Universal Robots PolyScope program: Weight_detection.urp

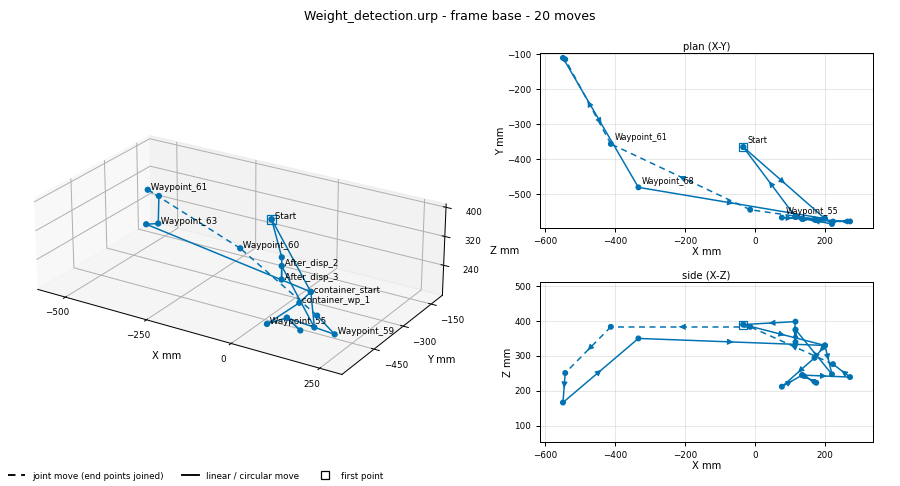
[picture p0: tool path of Weight_detection.urp in frame base, 20 of 20 moves have a stored position in this frame; points joined in program order, loops and branches not executed]
Program Weight_detection (installation=default directory=/programs/02 Main Routines createdIn=5.19.0 lastSavedIn=5.19.0 robotSerialNumber=20245590068)
Calibrated DH parameters: a=[0.00013, -0.03651, -0.389144, 0.000102, 0.000008, 0]; d=[0.162613, 192.230671, -179.915756, -12.181517, 0.099698, 0.099535]; alpha=[1.57038, 0.002205, 0.004138, 1.570804, -1.571025, 0]; deltaTheta=[-0.000001, 1.484886, 4.928506, -0.130209, 0, 0]
InitVariablesNode
Robot Program (runOnlyOnce=true)
  Folder powder dispensing variable init
    Start_thread := False
    kp := 0.0005
    ki := 0.002
    kd := 0.02
    dt := 0.05
    Weight_value := get_weight()
    Target_weight :=  (valueSource=Operator message=Enter the Target weight to be dispensed in gm valueType=Float)
    Integral_error := 0
    current_error := 0
    previous_error := 0
    tilt_increment := 0
    tilt_angle := -1
  Script file /programs/04 Scripts/Weight_scale_socket.script
    | def get_weight():
    | 	socket_open("192.168.12.190", 3002)
    | 	textmsg("socket opened successfully!")
    | 	socket_send_string("GET_WEIGHT")
    | 	sync()
    | 	sleep(0.5)
    | 	receiveFromServ = socket_read_ascii_float(6)
    | 	while (receiveFromServ[0] <1):
    | 		sleep(0.5)
    | 		receiveFromServ = socket_read_ascii_float(1)
    | 		textmsg("retrying read:", receiveFromServ)
    | 	end
    | 	textmsg("Received weight:", receiveFromServ[1])
    | 	socket_close()
    | 	return receiveFromServ[1]
    | end
  Script file /programs/04 Scripts/dosing_pid.script
    | def dosing_pid(Target_weight):
    | 	#kp = 0.005
    | 	#ki = 0.02
    | 	#kd = 0.2
    | 	#dt = 0.05
    | 	#current_error = 0.0
    | 	#Integral_error = 0.0
    | 	#previous_error = 0.0
    | 	#tilt_angle = -1.0
    | 	max_tilt_angle = -0.55
    | 	#current_pose = get_actual_tcp_pose()
    | 
    | 	while ( Weight_value < Target_weight and tilt_angle < max_tilt_angle):
    | 		Weight_value = get_weight()
    | 		current_error = Target_weight - Weight_value
    | 		Integral_error = Integral_error + current_error*dt
    | 		derivative = (current_error - previous_error) / dt
    | 		tilt_increment = (kp * current_error) + (ki * Integral_error) + (kd * derivative)
    | 		current_pose = get_actual_tcp_pose()
    | 		tilt_angle = current_pose[4]
    | 		new_pose = pose_trans(current_pose, p[(tilt_increment/5), 0, 0, 0, tilt_increment, 0])
    | 		movel(new_pose, a = 0.075, v = 0.025, t = 0, r = 0)
    | 		previous_error = current_error
    | 		sleep(dt)
    | 	end
    | end
  MoveL speed 250 mm/s, acceleration 1200 mm/s^2 (useActiveTCP=true) feature=Base
    Waypoint Start: TCP in base x=-33.065 y=-365.399 z=389.873 mm, rx=0 ry=0 rz=2.7258 rad; joints [-73.774, -70.638, -96.716, -102.629, 90.121, 40.001] deg; TCP offset x=0 y=0 z=161 mm, rx=3.1415 ry=0 rz=0 rad
  SuppressedNode
    MoveL speed 50 mm/s, acceleration 300 mm/s^2 (useActiveTCP=true) feature=Base
      Waypoint Waypoint_53: motionParameters(jointSpeed=1.047198 jointAcceleration=1.396263 cartesianSpeed=0.1 cartesianAcceleration=0.3); TCP in base x=200.65 y=-570.239 z=330.084 mm, rx=1.3605 ry=0.0217 rz=2.6816 rad; joints [-43.952, -124.342, -49.589, -141.868, 58.423, 68.107] deg
      Waypoint Waypoint_54: motionParameters(jointSpeed=1.047198 jointAcceleration=1.396263 cartesianSpeed=0.05 cartesianAcceleration=0.3); TCP in base x=170.614 y=-572.151 z=294.509 mm, rx=1.2595 ry=-0.0083 rz=2.7877 rad; joints [-46.577, -118.755, -62.143, -128.361, 58.907, 59.792] deg
      Loop Counting (count=3) loopVariable(name=Loop_4)
        Waypoint Waypoint_55: motionParameters(jointSpeed=1.047198 jointAcceleration=1.396263 cartesianSpeed=0.05 cartesianAcceleration=0.3); TCP in base x=77.281 y=-567.309 z=212.068 mm, rx=1.2595 ry=-0.0083 rz=2.7877 rad; joints [-52.608, -113.129, -83.31, -109.754, 55.252, 54.186] deg
          Until TOOL_CONTACT_DETECTION (allowActions=false retraction=0 decelerationAcceleration=3 decelerationAngularAcceleration=34.906585)
        Waypoint Waypoint_56: motionParameters(jointSpeed=1.047198 jointAcceleration=1.396263 cartesianSpeed=0.05 cartesianAcceleration=0.3); TCP in base x=135.568 y=-570.868 z=245.215 mm, rx=1.4769 ry=-0.0183 rz=2.6796 rad; joints [-47.325, -120.782, -69.397, -128.377, 54.155, 64.498] deg
      Loop Counting (count=2) loopVariable(name=Loop_5)
        Waypoint Waypoint_1: motionParameters(jointSpeed=1.047198 jointAcceleration=1.396263 cartesianSpeed=0.4 cartesianAcceleration=1.2); TCP in base x=175.61 y=-574.617 z=223.224 mm, rx=1.7438 ry=-0.031 rz=2.516 rad; joints [-43.942, -131.598, -59.719, -142.336, 52.9, 75.006] deg
        Waypoint Waypoint_56: motionParameters(jointSpeed=1.047198 jointAcceleration=1.396263 cartesianSpeed=0.05 cartesianAcceleration=0.3); TCP in base x=135.568 y=-570.868 z=245.215 mm, rx=1.4769 ry=-0.0183 rz=2.6796 rad; joints [-47.325, -120.782, -69.397, -128.377, 54.155, 64.498] deg
      Waypoint Waypoint_59: motionParameters(jointSpeed=1.047198 jointAcceleration=1.396263 cartesianSpeed=0.05 cartesianAcceleration=0.3); TCP in base x=272.401 y=-578.183 z=239.561 mm, rx=2.127 ry=0.1139 rz=2.1556 rad; joints [-37.816, -154.733, -25.502, -178.522, 53.445, 96.624] deg
      Waypoint Waypoint_58: motionParameters(jointSpeed=1.047198 jointAcceleration=1.396263 cartesianSpeed=0.05 cartesianAcceleration=0.3); TCP in base x=223.649 y=-578.478 z=276.546 mm, rx=2.1743 ry=-0.0441 rz=2.0587 rad; joints [-41.771, -153.265, -25.455, -184.54, 55.381, 96.631] deg
  SuppressedNode
    MoveJ speed 30 deg/s, acceleration 50 deg/s^2 (useActiveTCP=true) feature=Base
      Waypoint Waypoint_60: motionParameters(jointSpeed=0.349066 jointAcceleration=0.523599 cartesianSpeed=0.25 cartesianAcceleration=1.2 blendRadius=0.05); TCP in base x=-13.316 y=-544.772 z=383.372 mm, rx=2.2082 ry=0.0375 rz=2.0976 rad; joints [-53.447, -120.321, -68.514, -175.377, 39.556, 98.101] deg
      Waypoint Waypoint_61: motionParameters(jointSpeed=0.349066 jointAcceleration=0.523599 cartesianSpeed=0.25 cartesianAcceleration=1.2 blendRadius=0.05); TCP in base x=-412.189 y=-356.447 z=383.372 mm, rx=1.7517 ry=-0.74 rz=1.6007 rad; joints [-101.195, -120.321, -68.514, -175.377, 39.556, 98.101] deg
      Waypoint Waypoint_62: motionParameters(jointSpeed=0.349066 jointAcceleration=0.523599 cartesianSpeed=0.25 cartesianAcceleration=1.2); TCP in base x=-542.659 y=-114.282 z=251.262 mm, rx=1.813 ry=-0.6794 rz=1.6553 rad; joints [-123.661, -111.262, -103.952, -159.22, 12.548, 108.767] deg
  SuppressedNode
    MoveL speed 250 mm/s, acceleration 1200 mm/s^2 (useActiveTCP=true) feature=Base
      Waypoint Waypoint_63: motionParameters(jointSpeed=1.047198 jointAcceleration=1.396263 cartesianSpeed=0.05 cartesianAcceleration=0.3); TCP in base x=-532.496 y=-127.81 z=184.034 mm, rx=1.813 ry=-0.6794 rz=1.6553 rad; joints [-121.653, -117.001, -107.545, -147.984, 14.526, 106.805] deg
      If Target_weight<Weight_value (checkContinuously=true)
        Script: dosing_pid()
      Waypoint Waypoint_64: motionParameters(jointSpeed=1.047198 jointAcceleration=1.396263 cartesianSpeed=0.05 cartesianAcceleration=0.3); TCP in base x=-576.035 y=-66.27 z=306.74 mm, rx=0.8621 ry=-0.2554 rz=2.1952 rad; joints [-142.141, -87.685, -107.535, -64.498, 50.077, -8.596] deg
      Waypoint Waypoint_65: motionParameters(jointSpeed=1.047198 jointAcceleration=1.396263 cartesianSpeed=0.05 cartesianAcceleration=0.3); TCP in base x=-581.965 y=-59.291 z=312.082 mm, rx=0.8621 ry=-0.2554 rz=2.1952 rad; joints [-143.275, -88.018, -106.65, -64.116, 50.29, -10.05] deg
      Waypoint Waypoint_66: motionParameters(jointSpeed=1.047198 jointAcceleration=1.396263 cartesianSpeed=0.5 cartesianAcceleration=1.2); TCP in base x=-581.965 y=-59.291 z=290.576 mm, rx=0.8621 ry=-0.2554 rz=2.1952 rad; joints [-143.281, -88.87, -109.094, -60.824, 50.286, -10.043] deg
      Waypoint Waypoint_67: TCP in base x=-581.965 y=-59.291 z=350.142 mm, rx=1.7575 ry=-0.6778 rz=1.6965 rad; joints [-131.863, -101.687, -97.87, -162.913, 4.302, 96.426] deg
  SuppressedNode
    MoveJ speed 60 deg/s, acceleration 80 deg/s^2 (useActiveTCP=true) feature=Base
      Waypoint Waypoint_68: motionParameters(jointSpeed=1.047198 jointAcceleration=1.396263 cartesianSpeed=0.25 cartesianAcceleration=1.2); TCP in base x=-333.293 y=-480.744 z=350.142 mm, rx=2.2175 ry=0.1409 rz=2.2091 rad; joints [-82.414, -101.687, -97.87, -162.913, 4.302, 96.426] deg
  Folder powder dispensing
    Loop While (checkContinuously=false) expression=Weight_value<Target_weight
      MoveL speed 50 mm/s, acceleration 300 mm/s^2 (useActiveTCP=true) feature=Base
        Waypoint container_start: motionParameters(jointSpeed=1.047198 jointAcceleration=1.396263 cartesianSpeed=0.1 cartesianAcceleration=0.3); TCP in base x=200.65 y=-570.239 z=330.084 mm, rx=1.3605 ry=0.0217 rz=2.6816 rad; joints [-43.952, -124.342, -49.589, -141.868, 58.423, 68.107] deg
        Waypoint container_wp_1: motionParameters(jointSpeed=1.047198 jointAcceleration=1.396263 cartesianSpeed=0.05 cartesianAcceleration=0.3); TCP in base x=170.614 y=-572.151 z=294.509 mm, rx=1.2595 ry=-0.0083 rz=2.7877 rad; joints [-46.577, -118.755, -62.143, -128.361, 58.907, 59.792] deg
        Loop Counting (count=2) loopVariable(name=Loop_2)
          Waypoint Waypoint_55: motionParameters(jointSpeed=1.047198 jointAcceleration=1.396263 cartesianSpeed=0.07 cartesianAcceleration=0.5); TCP in base x=77.281 y=-567.309 z=212.068 mm, rx=1.2595 ry=-0.0083 rz=2.7877 rad; joints [-52.608, -113.129, -83.31, -109.754, 55.252, 54.186] deg
            Until TOOL_CONTACT_DETECTION (allowActions=false retraction=-0.005 decelerationAcceleration=0.3 decelerationAngularAcceleration=34.906585)
          Waypoint Waypoint_56: motionParameters(jointSpeed=1.047198 jointAcceleration=1.396263 cartesianSpeed=0.05 cartesianAcceleration=0.3); TCP in base x=135.568 y=-570.868 z=245.215 mm, rx=1.4769 ry=-0.0183 rz=2.6796 rad; joints [-47.325, -120.782, -69.397, -128.377, 54.155, 64.498] deg
        Loop Counting (count=1) loopVariable(name=Loop_6)
          Waypoint Waypoint_1: motionParameters(jointSpeed=1.047198 jointAcceleration=1.396263 cartesianSpeed=0.4 cartesianAcceleration=1.2); TCP in base x=175.61 y=-574.617 z=223.224 mm, rx=1.7438 ry=-0.031 rz=2.516 rad; joints [-43.942, -131.598, -59.719, -142.336, 52.9, 75.006] deg
          Waypoint Waypoint_56: motionParameters(jointSpeed=1.047198 jointAcceleration=1.396263 cartesianSpeed=0.05 cartesianAcceleration=0.3); TCP in base x=135.568 y=-570.868 z=245.215 mm, rx=1.4769 ry=-0.0183 rz=2.6796 rad; joints [-47.325, -120.782, -69.397, -128.377, 54.155, 64.498] deg
        Waypoint Waypoint_59: motionParameters(jointSpeed=1.047198 jointAcceleration=1.396263 cartesianSpeed=0.05 cartesianAcceleration=0.3); TCP in base x=272.401 y=-578.183 z=239.561 mm, rx=2.127 ry=0.1139 rz=2.1556 rad; joints [-37.816, -154.733, -25.502, -178.522, 53.445, 96.624] deg
        Waypoint Waypoint_58: motionParameters(jointSpeed=1.047198 jointAcceleration=1.396263 cartesianSpeed=0.05 cartesianAcceleration=0.3); TCP in base x=223.649 y=-578.478 z=276.546 mm, rx=2.1743 ry=-0.0441 rz=2.0587 rad; joints [-41.771, -153.265, -25.455, -184.54, 55.381, 96.631] deg
      MoveJ speed 30 deg/s, acceleration 50 deg/s^2 (useActiveTCP=true) feature=Base
        Waypoint Waypoint_60: motionParameters(jointSpeed=0.349066 jointAcceleration=0.523599 cartesianSpeed=0.25 cartesianAcceleration=1.2 blendRadius=0.05); TCP in base x=-13.316 y=-544.772 z=383.372 mm, rx=2.2082 ry=0.0375 rz=2.0976 rad; joints [-53.447, -120.321, -68.514, -175.377, 39.556, 98.101] deg
        Waypoint Waypoint_61: motionParameters(jointSpeed=0.349066 jointAcceleration=0.523599 cartesianSpeed=0.25 cartesianAcceleration=1.2 blendRadius=0.05); TCP in base x=-412.189 y=-356.447 z=383.372 mm, rx=1.7517 ry=-0.74 rz=1.6007 rad; joints [-101.195, -120.321, -68.514, -175.377, 39.556, 98.101] deg
        Waypoint Waypoint_62: motionParameters(jointSpeed=0.349066 jointAcceleration=0.523599 cartesianSpeed=0.25 cartesianAcceleration=1.2); TCP in base x=-542.659 y=-114.282 z=251.262 mm, rx=1.813 ry=-0.6794 rz=1.6553 rad; joints [-123.661, -111.262, -103.952, -159.22, 12.548, 108.767] deg
      MoveL speed 250 mm/s, acceleration 1200 mm/s^2 (useActiveTCP=true) feature=Base
        Waypoint Waypoint_63: motionParameters(jointSpeed=1.047198 jointAcceleration=1.396263 cartesianSpeed=0.05 cartesianAcceleration=0.3); TCP in base x=-549.161 y=-110.18 z=166.726 mm, rx=1.813 ry=-0.6794 rz=1.6553 rad; joints [-124.639, -119.53, -107.045, -149.088, 11.631, 110.027] deg
        Start_thread := True
        Wait Sleep waitTime=0.5
        Loop While (checkContinuously=true) expression=Weight_value≤Target_weight and tilt_angle≤-0.53
          current_error := Target_weight-Weight_value
          Integral_error := Integral_error+current_error*dt
          derivative := (current_error-previous_error)/dt
          tilt_increment := (kp*current_error)+(ki*Integral_error)+(kd*derivative)
          current_pose := get_actual_tcp_pose()
          tilt_angle := current_pose[4]
          tilt_pose := pose_trans(current_pose, p[(tilt_increment/5), 0, 0, 0, tilt_increment, 0])
          Script: movel(tilt_pose, a=0.025, v=0.015, r=0.00001)
          previous_error := current_error
          Wait Sleep waitTime=0.01
        Start_thread := False
        SuppressedNode
          Waypoint Waypoint_64: motionParameters(jointSpeed=1.047198 jointAcceleration=1.396263 cartesianSpeed=0.03 cartesianAcceleration=0.1 blendRadius=0.05); TCP in base x=-542.998 y=-117.021 z=221.977 mm, rx=1.8981 ry=-0.7227 rz=1.5827 rad; joints [-123.845, -120.87, -101.018, -172.406, 14.907, 127.864] deg
        Weight_value := get_weight()
        tilt_angle := -1
        Wait Sleep waitTime=0.5
      MoveL speed 250 mm/s, acceleration 1200 mm/s^2 (useActiveTCP=true) feature=Base
        Waypoint Waypoint_68: motionParameters(jointSpeed=0.436332 jointAcceleration=0.523599 cartesianSpeed=0.1 cartesianAcceleration=0.2 blendRadius=0.05); TCP in base x=-333.293 y=-480.744 z=350.142 mm, rx=2.2175 ry=0.1409 rz=2.2091 rad; joints [-82.414, -101.687, -97.87, -162.913, 4.302, 96.426] deg
        Waypoint Waypoint_3: motionParameters(jointSpeed=0.523599 jointAcceleration=0.698132 cartesianSpeed=0.1 cartesianAcceleration=0.4); TCP in base x=200.65 y=-570.239 z=330.084 mm, rx=2.1694 ry=-0.0462 rz=2.0859 rad; joints [-42.299, -146.843, -29.534, -185.935, 54.213, 95.41] deg
      Integral_error := 0
      current_error := 0
      previous_error := 0
    MoveL speed 250 mm/s, acceleration 1200 mm/s^2 (useActiveTCP=true) feature=Base
      Waypoint After_disp_1: motionParameters(jointSpeed=1.047198 jointAcceleration=1.396263 cartesianSpeed=0.1 cartesianAcceleration=0.4); TCP in base x=220.679 y=-585.611 z=247.463 mm, rx=2.1694 ry=-0.0462 rz=2.0859 rad; joints [-42.137, -153.398, -28.891, -180.007, 54.392, 95.38] deg
      Waypoint After_disp_2: motionParameters(jointSpeed=1.047198 jointAcceleration=1.396263 cartesianSpeed=0.06 cartesianAcceleration=0.4); TCP in base x=116.305 y=-565.093 z=375.554 mm, rx=0.6852 ry=0.0694 rz=2.9347 rad; joints [-54.743, -104.699, -66.451, -113.962, 68.291, 45.526] deg
      Waypoint After_disp_3: TCP in base x=116.305 y=-565.093 z=339.674 mm, rx=0.6852 ry=0.0694 rz=2.9347 rad; joints [-54.753, -104.143, -72.429, -108.545, 68.299, 45.538] deg
      Waypoint After_disp_4: TCP in base x=116.305 y=-565.093 z=398.258 mm, rx=0.6852 ry=0.0694 rz=2.9347 rad; joints [-54.737, -105.327, -62.27, -117.512, 68.285, 45.518] deg
      Waypoint Start: motionParameters(jointSpeed=1.047198 jointAcceleration=1.396263 cartesianSpeed=0.15 cartesianAcceleration=0.6); TCP in base x=-33.065 y=-365.399 z=389.873 mm, rx=0 ry=0 rz=2.7258 rad; joints [-73.774, -70.638, -96.716, -102.629, 90.121, 40.001] deg
      Popup Message (haltProgram=false message=Powder dispensed successfully... inputType=Text)
Thread Thread_1 (runOnlyOnce=false)
  If Start_thread≟ True
    Weight_value := get_weight()
    Wait Sleep waitTime=0.25
    Script: sync()
